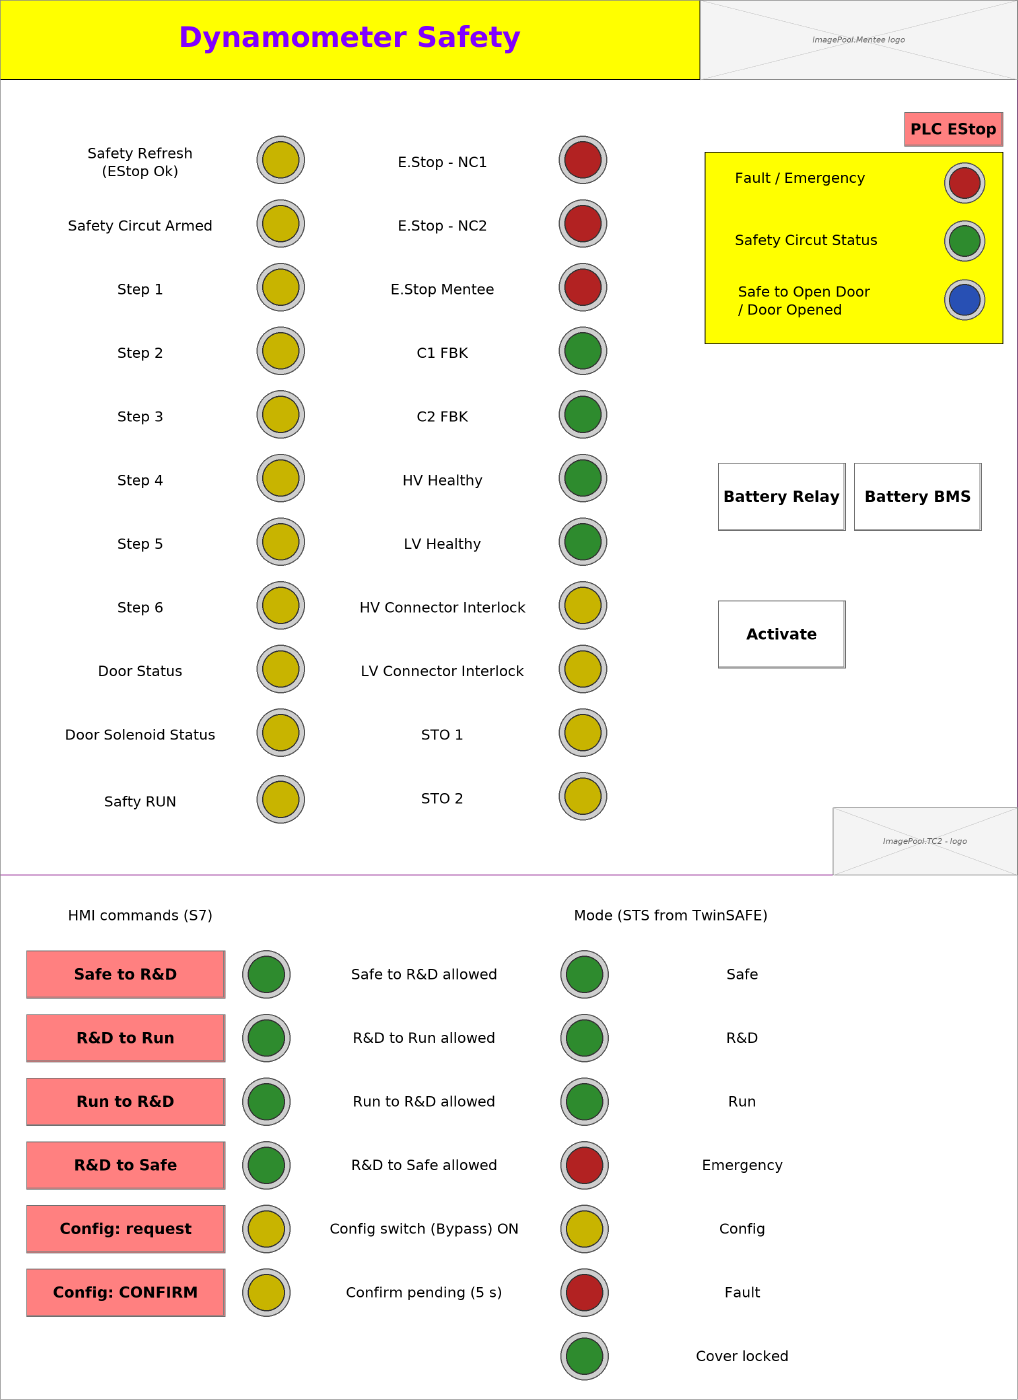
VISUALIZATION Visualization  // 1280x1760
    Rectangle (0,0 1280x1100)
    Rectangle (886,191 375x241)
    Rectangle (0,0 880x100)
    Lamp1 (318,166 70x70), variable: GVL_Safety.stTwinSAFE_IN.EStop_Ok, style: Lamp-Lamp1-Yellow
    Label (33,173 287x62), "Safety Refresh (EStop Ok)"
    Lamp1 (318,246 70x70), variable: GVL_Safety.stTwinSAFE_IN.Safety_Armed, style: Lamp-Lamp1-Yellow
    Label (33,253 287x62), "Safety Circut Armed"
    Lamp1 (318,326 70x70), variable: GVL_Safety.stTwinSAFE_IN.Speps.step1, style: Lamp-Lamp1-Yellow
    Label (33,333 287x62), "Step 1"
    Lamp1 (318,406 70x70), variable: GVL_Safety.stTwinSAFE_IN.Speps.step2, style: Lamp-Lamp1-Yellow
    Label (33,413 287x62), "Step 2"
    Lamp1 (318,486 70x70), variable: GVL_Safety.stTwinSAFE_IN.Speps.step3, style: Lamp-Lamp1-Yellow
    Label (33,493 287x62), "Step 3"
    Lamp1 (318,566 70x70), variable: GVL_Safety.stTwinSAFE_IN.Speps.step4, style: Lamp-Lamp1-Yellow
    Label (33,573 287x62), "Step 4"
    Lamp1 (318,646 70x70), variable: GVL_Safety.stTwinSAFE_IN.Speps.step5, style: Lamp-Lamp1-Yellow
    Label (33,653 287x62), "Step 5"
    Lamp1 (318,726 70x70), variable: GVL_Safety.stTwinSAFE_IN.Speps.step6, style: Lamp-Lamp1-Yellow
    Label (33,733 287x62), "Step 6"
    Lamp1 (318,806 70x70), variable: GVL_Safety.DoorMonitorFromPLC, style: Lamp-Lamp1-Yellow
    Label (33,813 287x62), "Door Status"
    Lamp1 (318,970 70x70), variable: GVL_Safety.stTwinSAFE_OUT.RUN, style: Lamp-Lamp1-Yellow
    Label (33,977 287x62), "Safty RUN"
    Lamp1 (318,886 70x70), variable: GVL_Safety.SolonoidStatus, style: Lamp-Lamp1-Yellow
    Label (33,893 287x62), "Door Solenoid Status"
    Button (1137,141 124x43), "PLC EStop", colour toggle: GVL_Safety.stTwinSAFE_OUT.EstopPLC
        toggle GVL_Safety.stTwinSAFE_OUT.EstopPLC
    Button (903,582 160x85), "Battery Relay", colour toggle: GVL_Safety.stTwinSAFE_OUT.BatRelay_CMD
        toggle GVL_Safety.stTwinSAFE_OUT.BatRelay_CMD
    Button (1074,582 160x85), "Battery BMS", colour toggle: GVL_Safety.stTwinSAFE_OUT.BatBMS_Cmd
        toggle GVL_Safety.stTwinSAFE_OUT.BatBMS_Cmd
    Lamp1 (698,166 70x70), variable: GVL_Safety.stTwinSAFE_IN.EStop_NC1, style: Lamp-Lamp1-Red
    Label (413,173 287x62), "E.Stop - NC1"
    Lamp1 (698,246 70x70), variable: GVL_Safety.stTwinSAFE_IN.EStop_NC2, style: Lamp-Lamp1-Red
    Label (413,253 287x62), "E.Stop - NC2"
    Lamp1 (698,326 70x70), variable: GVL_Safety.stTwinSAFE_IN.EStop_MantiRob, style: Lamp-Lamp1-Red
    Label (413,333 287x62), "E.Stop Mentee"
    Lamp1 (698,406 70x70), variable: GVL_Safety.stTwinSAFE_IN.C1_FBK, style: Lamp-Lamp1-Green
    Label (413,413 287x62), "C1 FBK"
    Lamp1 (698,486 70x70), variable: GVL_Safety.stTwinSAFE_IN.C2_FBK, style: Lamp-Lamp1-Green
    Label (413,493 287x62), "C2 FBK"
    Lamp1 (698,566 70x70), variable: GVL_Safety.stTwinSAFE_IN.HV_Healthy, style: Lamp-Lamp1-Green
    Label (413,573 287x62), "HV Healthy"
    Lamp1 (698,646 70x70), variable: GVL_Safety.stTwinSAFE_IN.LV_Healthy, style: Lamp-Lamp1-Green
    Label (413,653 287x62), "LV Healthy"
    Lamp1 (698,726 70x70), variable: GVL_Safety.stTwinSAFE_IN.HV_Interlock, style: Lamp-Lamp1-Yellow
    Label (413,733 287x62), "HV Connector Interlock"
    Lamp1 (698,806 70x70), variable: GVL_Safety.stTwinSAFE_IN.LV_Interlock, style: Lamp-Lamp1-Yellow
    Label (413,813 287x62), "LV Connector Interlock"
    Lamp1 (698,886 70x70), variable: GVL_Safety.stTwinSAFE_IN.STO_1, style: Lamp-Lamp1-Yellow
    Label (413,893 287x62), "STO 1"
    Lamp1 (698,966 70x70), variable: GVL_Safety.stTwinSAFE_IN.STO_2, style: Lamp-Lamp1-Yellow
    Label (413,973 287x62), "STO 2"
    Button (903,755 160x85), "Activate", colour toggle: GVL_IO.b_MotorCooling
        toggle GVL_IO.b_MotorCooling
    Image (880,0 400x100), image: ImagePool.Mentee logo
    Label (0,0 880x93), "Dynamometer Safety"
    Lamp1 (1183,200 60x60), variable: GVL_IO.RedLED, style: Lamp-Lamp1-Red
    Lamp1 (1183,273 60x60), variable: GVL_IO.GreenLED, style: Lamp-Lamp1-Green
    Lamp1 (1183,347 60x60), variable: GVL_IO.BlueLED, style: Lamp-Lamp1-Blue
    Label (921,193 195x62), "Fault / Emergency"
    Label (921,271 252x62), "Safety Circut Status"
    Label (925,347 252x62), "Safe to Open Door / Door Opened"
    Label (895,517 252x62), "Battery Control"
    Label (903,691 252x62), "Motor Cooling"
    Label (886,133 300x62), "System Status"
    Image (1047,1015 233x85), image: ImagePool.TC2 - logo
    Label (33,1120 287x62), "HMI commands (S7)"
    Label (700,1120 287x62), "Mode (STS from TwinSAFE)"
    Button (33,1195 250x60), "Safe to R&D", colour toggle: MAIN.bHmi_SafeToRnD
        toggle MAIN.bHmi_SafeToRnD
    Lamp1 (300,1190 70x70), variable: MAIN.bEn_SafeToRnD, style: Lamp-Lamp1-Green
    Label (390,1194 287x62), "Safe to R&D allowed"
    Button (33,1275 250x60), "R&D to Run", colour toggle: MAIN.bHmi_RnDToRun
        toggle MAIN.bHmi_RnDToRun
    Lamp1 (300,1270 70x70), variable: MAIN.bEn_RnDToRun, style: Lamp-Lamp1-Green
    Label (390,1274 287x62), "R&D to Run allowed"
    Button (33,1355 250x60), "Run to R&D", colour toggle: MAIN.bHmi_RunToRnD
        toggle MAIN.bHmi_RunToRnD
    Lamp1 (300,1350 70x70), variable: MAIN.bEn_RunToRnD, style: Lamp-Lamp1-Green
    Label (390,1354 287x62), "Run to R&D allowed"
    Button (33,1435 250x60), "R&D to Safe", colour toggle: MAIN.bHmi_RnDToSafe
        toggle MAIN.bHmi_RnDToSafe
    Lamp1 (300,1430 70x70), variable: MAIN.bEn_RnDToSafe, style: Lamp-Lamp1-Green
    Label (390,1434 287x62), "R&D to Safe allowed"
    Button (33,1515 250x60), "Config: request", colour toggle: MAIN.bHmi_CfgReq
        toggle MAIN.bHmi_CfgReq
    Lamp1 (300,1510 70x70), variable: GVL_Safety.stTwinSAFE_OUT.Bypass_C1C2, style: Lamp-Lamp1-Yellow
    Label (390,1514 287x62), "Config switch (Bypass) ON"
    Button (33,1595 250x60), "Config: CONFIRM", colour toggle: MAIN.bHmi_CfgConfirm
        toggle MAIN.bHmi_CfgConfirm
    Lamp1 (300,1590 70x70), variable: MAIN.bCfgPending, style: Lamp-Lamp1-Yellow
    Label (390,1594 287x62), "Confirm pending (5 s)"
    Lamp1 (700,1190 70x70), variable: GVL_Safety.stTwinSAFE_IN.STS_SAFE, style: Lamp-Lamp1-Green
    Label (790,1194 287x62), "Safe"
    Lamp1 (700,1270 70x70), variable: GVL_Safety.stTwinSAFE_IN.STS_RND, style: Lamp-Lamp1-Green
    Label (790,1274 287x62), "R&D"
    Lamp1 (700,1350 70x70), variable: GVL_Safety.stTwinSAFE_IN.STS_RUN, style: Lamp-Lamp1-Green
    Label (790,1354 287x62), "Run"
    Lamp1 (700,1430 70x70), variable: GVL_Safety.stTwinSAFE_IN.STS_EMG, style: Lamp-Lamp1-Red
    Label (790,1434 287x62), "Emergency"
    Lamp1 (700,1510 70x70), variable: GVL_Safety.stTwinSAFE_IN.STS_CFG, style: Lamp-Lamp1-Yellow
    Label (790,1514 287x62), "Config"
    Lamp1 (700,1590 70x70), variable: GVL_Safety.stTwinSAFE_IN.STS_FAULT, style: Lamp-Lamp1-Red
    Label (790,1594 287x62), "Fault"
    Lamp1 (700,1670 70x70), variable: GVL_Safety.stTwinSAFE_IN.STS_COVER_LOCKED, style: Lamp-Lamp1-Green
    Label (790,1674 287x62), "Cover locked"
END_VISUALIZATION

(* stored: Version 1.1.0.1, ProductVersion 3.1.4026.18
   Visu Visualization: Id {7277df54-efcd-437b-8c25-efbbf80b43b5} *)
